// Mock of the mirror covers (I_MirrorCovers): Open/Close take effect at once, unless bHoldClose is set: then Close is only counted
// and the covers stay open until the test sets bClosed (a slow closing, IAG50cm#187).
FUNCTION_BLOCK FB_CoversMock IMPLEMENTS BROTLib.I_MirrorCovers
VAR
	bOpened		: BOOL;
	bClosed		: BOOL := TRUE;
	bFailed		: BOOL;
	bHoldClose	: BOOL;
	nOpenCalls	: UINT;
	nCloseCalls	: UINT;
END_VAR

METHOD Open : BOOL
bOpened := TRUE;
bClosed := FALSE;
nOpenCalls := nOpenCalls + 1;
Open := TRUE;
END_METHOD

METHOD Close : BOOL
bOpened := FALSE;
IF NOT bHoldClose THEN
	bClosed := TRUE;
END_IF
nCloseCalls := nCloseCalls + 1;
Close := TRUE;
END_METHOD

// while bHold is TRUE a Close() is only counted and the covers stay open (a slow closing, IAG50cm#187)
METHOD HoldClose
VAR_INPUT
	bHold	: BOOL;
END_VAR
bHoldClose := bHold;
END_METHOD

// the held closing is done: the covers are closed now
METHOD FinishClose
bHoldClose := FALSE;
bOpened := FALSE;
bClosed := TRUE;
END_METHOD

METHOD Reset : BOOL
bFailed := FALSE;
Reset := TRUE;
END_METHOD

PROPERTY Opened : BOOL
GET
Opened := bOpened;
END_GET
END_PROPERTY

PROPERTY Closed : BOOL
GET
Closed := bClosed;
END_GET
END_PROPERTY

PROPERTY Error : BOOL
GET
Error := bFailed;
END_GET
END_PROPERTY

END_FUNCTION_BLOCK

(* stored: Version 1.1.0.1, ProductVersion 3.1.4024.15
   POU FB_CoversMock: Id {012aa109-a307-4f4a-912d-8723ceeda833}, SpecialFunc None
   Method Open: Id {13845e21-9c3e-4dac-b959-05571002f911}
   Method Close: Id {656096ac-ec16-41d0-b289-34747ce3f99b}
   Method HoldClose: Id {d7d1cc71-70fb-451a-98a6-0959d77f9320}
   Method FinishClose: Id {6550a56f-c343-4224-a85a-2f5a08bdcf22}
   Method Reset: Id {4ff33918-9b37-404a-9749-6f3afb8baa3c}
   Property Opened: Id {fba570be-a0a2-4e23-9865-61e4da490848}
   Get Get: Id {d58103d1-991b-4192-8a45-f3aa4cebda72}
   Property Closed: Id {7625856f-be1f-47bf-b814-ccb6a41d741b}
   Get Get: Id {d7e43db7-68e3-4543-9de8-f14deb00cbeb}
   Property Error: Id {a5ed7b97-9402-4c8f-9ba4-5e6a096dcc20}
   Get Get: Id {e0c06a2c-4379-42ec-b938-ee5f2578c49c} *)
